VAR_GLOBAL
    bUpperButton : BOOL;
    bLowerButton : BOOL;
    bOuterSpotsRelay : BOOL;
    bMiddleSpotRelay : BOOL;
END_VAR

(* stored: Version 1.1.0.1
   GVL GVL_HallSimulation: Id {818a25ce-54ac-4fc2-a2ef-5916ec994a4d} *)
